(*
SPDX-FileCopyrightText: c 2026 Oleksandr Tiutyk <trofimich@gmail.com>
SPDX-License-Identifier: MIT
License: https://opensource.org/license/mit
*)

(*!
<summary>Checks matching and missing keys with raw and borrowed generic queries.</summary>
<description>
Borrows one group-owned dictionary reserved for this case. Use from one task at a stable address.
Teardown clears entries owned by the dictionary before publication.
</description>
*)

{attribute 'no_assign'}
{attribute 'no_explicit_call' := 'do not call this function block directly'}
FUNCTION_BLOCK DictionaryContainsTest EXTENDS TOF_Testing.SingleCycleTest
VAR_STAT
	{attribute 'hide'}
	_ClassName : STRING := __POUNAME();
END_VAR
VAR
	_Dictionary : TOF_Collections.IDictionary;
END_VAR

(*!
<summary>Clears the fixture before the runner publishes the result.</summary>
<description>
Also runs after an unexpected exception interrupts the case.
</description>
*)
METHOD PROTECTED AfterTest
_Dictionary.Clear();
END_METHOD

//! <summary>Borrows the concrete class name. Callers must not modify it.</summary>
{attribute 'monitoring' := 'call'}
PROPERTY ClassName : REFERENCE TO STRING
GET
ClassName REF= _ClassName;
END_GET
END_PROPERTY

(*!
<summary>Checks matching and missing keys with raw and borrowed generic queries.</summary>
*)
METHOD PROTECTED ExecuteTest
VAR
	keys : ARRAY [0..6] OF INT := [0, 1, 2, 3, 4, 5, 6];
	values : ARRAY [0..6] OF STRING :=
		['String0', 'String1', 'String2', 'String3', 'String4', 'String5', 'String6'];
	i : DINT;
	missingKey : INT := 9;
	query : TOF_Core.GENERIC_VALUE;
END_VAR
FOR i := 6 TO 0 BY -1 DO
	_Dictionary.SetCopy(key := keys[i], value := values[i]);
END_FOR

_Dictionary.SetCopy(key := keys[3], value := values[3]);

Assert.ThatBool(
	actual := _Dictionary.ContainsKey(key := keys[3]),
	message := "ContainsKey must find the stored key"
).IsTrue();

Assert.ThatBool(
	actual := _Dictionary.ContainsKey(key := missingKey),
	message := "ContainsKey must reject an absent key"
).IsFalse();

query := TOF_Core.GenericValueFactory.FromIntReference(value := keys[3]);
Assert.ThatBool(
	actual := _Dictionary.ContainsGenericKey(key := query, releaseKey := FALSE),
	message := "ContainsGenericKey must find the stored key"
).IsTrue();

query := TOF_Core.GenericValueFactory.FromIntReference(value := missingKey);
Assert.ThatBool(
	actual := _Dictionary.ContainsGenericKey(key := query, releaseKey := FALSE),
	message := "ContainsGenericKey must reject an absent key"
).IsFalse();

Assert.ThatDInt(
	actual := _Dictionary.Length,
	message := "Lookup must preserve all seven entries"
).ToBe(expected := DINT#7);
END_METHOD

(*!
<summary>Binds the dictionary fixture for this case.</summary>
<description>
Stores a borrowed interface without invoking the fixture. The owning group keeps it alive and
reserves it for this case. TestElement initializes the name and parent.
</description>
<param name="name">Display name of this case.</param>
<param name="parent">Group that owns this case.</param>
<param name="dictionary">Required live dictionary reserved for this case.</param>
*)
METHOD FB_init : BOOL
VAR_INPUT
	bInitRetains: BOOL; // TRUE: the retain variables are initialized (reset warm / reset cold)
	bInCopyCode: BOOL; // TRUE: the instance will be copied to the copy code afterward (online change)
	name : WSTRING;
	parent : TOF_Testing.ITestElement;
	dictionary : TOF_Collections.IDictionary;
END_VAR
_Dictionary := dictionary;
FB_init := TRUE;
END_METHOD

//! <summary>Borrows the compiler-initialized namespace name. Callers must not modify it.</summary>
{attribute 'monitoring' := 'call'}
PROPERTY NamespaceName : REFERENCE TO STRING
GET
NamespaceName REF= CurrentNamespace.Name;
END_GET
END_PROPERTY

//! <summary>Reports the concrete instance size in bytes.</summary>
{attribute 'monitoring' := 'call'}
PROPERTY SelfSize : ULINT
GET
SelfSize := XSIZEOF(THIS^);
END_GET
END_PROPERTY

END_FUNCTION_BLOCK

(* stored: Version 1.1.0.1, ProductVersion 3.1.4026.21
   POU DictionaryContainsTest: Id {2d7a40c9-cbba-45f4-ba83-476cbde093c0}, SpecialFunc None
   Method AfterTest: Id {cf996799-1669-4115-b0d5-304f335c59ba}
   Property ClassName: Id {cc3a92c8-6716-4aa2-b93f-62e4ba12463f}
   Get Get: Id {ce07f8d2-dbf3-401c-9390-2a45f7b05a3f}
   Method ExecuteTest: Id {953a4708-e6c0-4c93-8d3b-3f7d058a91ff}
   Method FB_init: Id {f8304e8b-650e-4a5d-b552-76f39363504b}
   Property NamespaceName: Id {715962f3-c34b-4f8f-a738-5da52b32941e}
   Get Get: Id {fa995312-0b65-4c06-91e0-97d44e7f9b81}
   Property SelfSize: Id {e3e510d7-9e34-4923-a36b-b8f6974ad375}
   Get Get: Id {ebc8ef7f-452b-473c-b764-6c70c4737628} *)
